INTERFACE ITcoState EXTENDS ITcoObject, ITcoRestorable

PROPERTY IsAutoRestoreEnabled : BOOL
GET
END_GET
END_PROPERTY

PROPERTY LastStateChangeCycle : ULINT
GET
END_GET
END_PROPERTY

METHOD RestoreObject : ITcoObjectRestorer
VAR_INPUT
	Obj : ITcoRestorable;
END_VAR
END_METHOD

PROPERTY State : INT
GET
END_GET
END_PROPERTY

END_INTERFACE

(* stored: Version 1.1.0.1
   Itf ITcoState: Id {c649817a-92de-4bd9-bb87-c0d72fad7509}
   Property IsAutoRestoreEnabled: Id {919401ee-55fe-4554-8ddf-1a407786ef18}
   Get Get: Id {87b763ca-6a82-43eb-8730-8dd9412bbc83}
   Property LastStateChangeCycle: Id {92216c9b-4911-48a2-a6ff-b6246c33da8c}
   Get Get: Id {78ddabb3-69a5-4bb1-a9d6-f1af6af00fdd}
   Method RestoreObject: Id {4a8a2884-a04a-427f-a212-93f7d99ca614}
   Property State: Id {ffa51ee9-dcc1-48dd-ac68-d06a65059caf}
   Get Get: Id {b970a776-b81b-430c-827a-7496827f2909} *)
